ABB RAPID module: TopSurf.mod

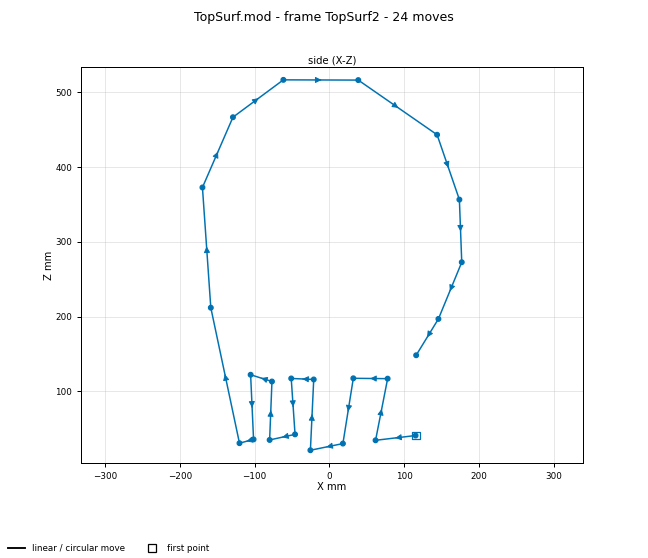
[picture p0: tool path of TopSurf.mod in frame TopSurf2, 24 of 27 moves have a stored position in this frame; points joined in program order, loops and branches not executed]
%%%
  VERSION:1
  LANGUAGE:ENGLISH
%%%
MODULE MOD_TopSurf

    ! -------------------------------
    ! Define customized variables here
    ! ...

	! Tool variables:
	PERS tooldata ToolRDK2 := [TRUE,[[-397.000,-4.578,191.692],[0.70710678,0.00000000,-0.70710678,0.00000001]],[1,[0,0,20],[1,0,0,0],0,0,0.005]];

	! Reference variables:
	PERS wobjdata TopSurf2 := [FALSE, TRUE, "", [[0,0,0],[1,0,0,0]],[[1336.130,0.000,735.410],[0.50000000,0.50000000,0.50000000,0.50000000]]];

	PROC TT0deg()
		ConfJ \On;
		ConfL \Off;
		MoveAbsJ [[0.000000,0.000000,0.000000,0.000000,0.000000,0.000000],[9E+09,9E+09,9E+09,9E+09,9E+09,9E+09]],v500,z1,ToolRDK2 \WObj:=TopSurf2;
	ENDPROC

	PROC Main()
		ConfJ \On;
		ConfL \Off;
		! Program generated by VerticalBot Studio for ABB IRB 2600-12/1.85 on 25/10/2026 12:00:00
		! Using nominal kinematics.
		TT0deg;
		TopSurf2 := [FALSE, TRUE, "", [[0,0,0],[1,0,0,0]],[[1336.130,0.000,735.410],[0.50000000,0.50000000,0.50000000,0.50000000]]];
		ToolRDK2 := [TRUE,[[-397.000,-4.578,191.692],[0.70710678,0.00000000,-0.70710678,0.00000001]],[1,[0,0,20],[1,0,0,0],0,0,0.005]];
		MoveAbsJ [[-2.762230,35.281600,-32.244600,94.063100,36.825000,84.928900],[9E+09,9E+09,9E+09,9E+09,9E+09,9E+09]],v500,z1,ToolRDK2 \WObj:=TopSurf2;
		MoveAbsJ [[3.888270,37.649400,-27.622300,84.244200,-60.438300,101.547000],[9E+09,9E+09,9E+09,9E+09,9E+09,9E+09]],v500,z1,ToolRDK2 \WObj:=TopSurf2;
		GunOn 1;
		MoveL [[115.290,-0.000,40.893],[0.66951661,0.66951663,0.22748073,-0.22748077],[-1,1,1,2],[9E+09,9E+09,9E+09,9E+09,9E+09,9E+09]],v500,z1,ToolRDK2 \WObj:=TopSurf2;
		MoveL [[61.769,-0.000,34.498],[0.66824739,0.66824741,0.23118262,-0.23118267],[0,0,1,1],[9E+09,9E+09,9E+09,9E+09,9E+09,9E+09]],v500,z1,ToolRDK2 \WObj:=TopSurf2;
		MoveL [[77.918,0.000,116.954],[0.67411479,0.67411479,0.21346957,-0.21346957],[0,0,1,1],[9E+09,9E+09,9E+09,9E+09,9E+09,9E+09]],v500,z1,ToolRDK2 \WObj:=TopSurf2;
		MoveL [[32.029,0.000,117.425],[0.67416339,0.67416339,0.21331602,-0.21331602],[0,0,1,1],[9E+09,9E+09,9E+09,9E+09,9E+09,9E+09]],v500,z1,ToolRDK2 \WObj:=TopSurf2;
		MoveL [[18.094,-0.000,30.124],[0.66795555,0.66795555,0.23202454,-0.23202454],[0,0,1,1],[9E+09,9E+09,9E+09,9E+09,9E+09,9E+09]],v500,z1,ToolRDK2 \WObj:=TopSurf2;
		MoveL [[-25.377,-0.000,21.201],[0.66687834,0.66687834,0.23510269,-0.23510270],[0,0,1,1],[9E+09,9E+09,9E+09,9E+09,9E+09,9E+09]],v500,z1,ToolRDK2 \WObj:=TopSurf2;
		MoveL [[-20.929,0.000,115.878],[0.67369753,0.67369752,0.21478279,-0.21478278],[0,0,1,1],[9E+09,9E+09,9E+09,9E+09,9E+09,9E+09]],v500,z1,ToolRDK2 \WObj:=TopSurf2;
		MoveL [[-51.029,0.000,117.232],[0.67365028,0.67365028,0.21493093,-0.21493093],[0,0,1,1],[9E+09,9E+09,9E+09,9E+09,9E+09,9E+09]],v500,z1,ToolRDK2 \WObj:=TopSurf2;
		MoveL [[-45.916,-0.000,42.441],[0.66826232,0.66826233,0.23113949,-0.23113950],[0,0,1,1],[9E+09,9E+09,9E+09,9E+09,9E+09,9E+09]],v500,z1,ToolRDK2 \WObj:=TopSurf2;
		MoveL [[-79.907,-0.000,34.972],[0.66736193,0.66736194,0.23372644,-0.23372644],[0,0,1,1],[9E+09,9E+09,9E+09,9E+09,9E+09,9E+09]],v500,z1,ToolRDK2 \WObj:=TopSurf2;
		MoveL [[-76.800,0.000,113.142],[0.67321469,0.67321469,0.21629141,-0.21629141],[0,0,1,1],[9E+09,9E+09,9E+09,9E+09,9E+09,9E+09]],v500,z1,ToolRDK2 \WObj:=TopSurf2;
		MoveL [[-105.332,0.000,122.191],[0.67370783,0.67370783,0.21475045,-0.21475045],[0,0,1,1],[9E+09,9E+09,9E+09,9E+09,9E+09,9E+09]],v500,z1,ToolRDK2 \WObj:=TopSurf2;
		MoveL [[-101.402,-0.000,35.713],[0.66719553,0.66719554,0.23420101,-0.23420104],[0,0,1,1],[9E+09,9E+09,9E+09,9E+09,9E+09,9E+09]],v500,z1,ToolRDK2 \WObj:=TopSurf2;
		MoveL [[-120.231,-0.000,30.646],[0.66659020,0.66659020,0.23591842,-0.23591844],[0,0,1,1],[9E+09,9E+09,9E+09,9E+09,9E+09,9E+09]],v500,z1,ToolRDK2 \WObj:=TopSurf2;
		MoveL [[-158.578,-0.000,211.837],[0.67989399,0.67989399,0.19427858,-0.19427858],[0,2,-1,0],[9E+09,9E+09,9E+09,9E+09,9E+09,9E+09]],v500,z1,ToolRDK2 \WObj:=TopSurf2;
		MoveL [[-169.769,-0.000,372.687],[0.68989069,0.68989069,0.15508330,-0.15508330],[0,2,-1,0],[9E+09,9E+09,9E+09,9E+09,9E+09,9E+09]],v500,z1,ToolRDK2 \WObj:=TopSurf2;
		MoveL [[-128.964,0.000,466.626],[0.69493868,0.69493868,0.13061485,-0.13061485],[0,2,-1,0],[9E+09,9E+09,9E+09,9E+09,9E+09,9E+09]],v500,z1,ToolRDK2 \WObj:=TopSurf2;
		MoveL [[-61.529,0.000,516.598],[0.69594843,0.69594843,0.12512308,-0.12512308],[0,2,-1,0],[9E+09,9E+09,9E+09,9E+09,9E+09,9E+09]],v500,z1,ToolRDK2 \WObj:=TopSurf2;
		MoveL [[38.647,0.000,516.273],[0.69521781,0.69521781,0.12912086,-0.12912086],[0,2,-1,0],[9E+09,9E+09,9E+09,9E+09,9E+09,9E+09]],v500,z1,ToolRDK2 \WObj:=TopSurf2;
		MoveL [[144.073,0.000,443.157],[0.69160511,0.69160511,0.14724934,-0.14724934],[0,0,1,1],[9E+09,9E+09,9E+09,9E+09,9E+09,9E+09]],v500,z1,ToolRDK2 \WObj:=TopSurf2;
		MoveL [[173.888,-0.000,356.448],[0.68759917,0.68759917,0.16494659,-0.16494659],[0,0,1,1],[9E+09,9E+09,9E+09,9E+09,9E+09,9E+09]],v500,z1,ToolRDK2 \WObj:=TopSurf2;
		MoveL [[177.057,0.000,272.670],[0.68344550,0.68344550,0.18138976,-0.18138976],[0,0,1,1],[9E+09,9E+09,9E+09,9E+09,9E+09,9E+09]],v500,z1,ToolRDK2 \WObj:=TopSurf2;
		MoveL [[145.838,-0.000,196.841],[0.67931130,0.67931130,0.19630627,-0.19630627],[0,0,1,1],[9E+09,9E+09,9E+09,9E+09,9E+09,9E+09]],v500,z1,ToolRDK2 \WObj:=TopSurf2;
		GunOn 0;
		MoveL [[116.077,0.000,148.259],[0.67637750,0.67637750,0.20618797,-0.20618797],[0,0,1,1],[9E+09,9E+09,9E+09,9E+09,9E+09,9E+09]],v500,z1,ToolRDK2 \WObj:=TopSurf2;
	ENDPROC

ENDMODULE
